(* IEC 61131-3 sources: llm-plc-st-eval/data/processed_definitivo/qwen2.5-coder_14b/C7/few_shot, 3 files *)

(* ---- ejec_1.st ---- *)
FUNCTION_BLOCK FB_Contador
VAR_INPUT
    sensorPieza : BOOL; (* Contacto NA que alimenta CU *)
    btnReset : BOOL; (* Contacto NA que alimenta RESET *)
END_VAR
VAR_OUTPUT
    loteListo : BOOL; (* Bobina que se activa cuando C1.Q es TRUE *)
    cuenta : INT; (* Valor actual del contador *)
END_VAR
VAR
    C1 : CTU; (* Contador ascendente *)
END_VAR

(* Configuración del contador *)
C1.PV := 12; (* Valor preestablecido a 12 *)

(* Rama 1: alimentar CU y RESET *)
IF sensorPieza THEN
    C1.CU := TRUE;
ELSE
    C1.CU := FALSE;
END_IF

IF btnReset THEN
    C1.RESET := TRUE;
ELSE
    C1.RESET := FALSE;
END_IF

(* Rama 2: alimentar loteListo *)
loteListo := C1.Q;

(* Rama 3: transferir C1.CV a cuenta *)
cuenta := C1.CV;

(* Actualizar el contador *)
C1();

END_FUNCTION_BLOCK

(* ---- ejec_2.st ---- *)
FUNCTION_BLOCK FB_Contador
VAR_INPUT
    sensorPieza : BOOL; (* Contacto NA que alimenta CU *)
    btnReset : BOOL; (* Contacto NA que alimenta RESET *)
END_VAR
VAR_OUTPUT
    loteListo : BOOL; (* Bobina que se activa cuando C1.Q es TRUE *)
    cuenta : INT; (* Valor actual del contador *)
END_VAR
VAR
    C1 : CTU; (* Contador ascendente *)
END_VAR

(* Configuración del contador *)
C1.PV := 12; (* Valor preestablecido del contador *)

(* Rama 1: alimentar CU y RESET *)
IF sensorPieza THEN
    C1.CU := TRUE;
ELSE
    C1.CU := FALSE;
END_IF

IF btnReset THEN
    C1.RESET := TRUE;
ELSE
    C1.RESET := FALSE;
END_IF

(* Rama 2: alimentar loteListo *)
loteListo := C1.Q;

(* Rama 3: transferir C1.CV a cuenta *)
cuenta := C1.CV;

(* Ejecutar el contador *)
C1();

END_FUNCTION_BLOCK

(* ---- ejec_3.st ---- *)
FUNCTION_BLOCK FB_Contador
VAR_INPUT
    sensorPieza : BOOL; (* Contacto NA para contar *)
    btnReset : BOOL; (* Contacto NA para resetear el contador *)
END_VAR
VAR_OUTPUT
    loteListo : BOOL; (* Bobina que se activa cuando se alcanza el lote *)
    cuenta : INT; (* Valor actual del contador *)
END_VAR
VAR
    C1 : CTU; (* Contador ascendente *)
END_VAR

(* Configuración del contador *)
C1.PV := 12; (* Valor preestablecido del contador *)

(* Rama 1: Conteo *)
IF sensorPieza THEN
    C1.CU := TRUE; (* Incrementa el contador *)
ELSE
    C1.CU := FALSE;
END_IF

(* Rama 2: Reset *)
IF btnReset THEN
    C1.RESET := TRUE; (* Resetea el contador *)
ELSE
    C1.RESET := FALSE;
END_IF

(* Rama 3: Actualización del contador *)
C1(); (* Ejecuta el contador *)
cuenta := C1.CV; (* Transfiere el valor actual del contador a la variable cuenta *)

(* Rama 4: Lote listo *)
loteListo := C1.Q; (* La bobina se activa cuando se alcanza el valor preestablecido *)
END_FUNCTION_BLOCK
